// Liaison d'un résultat (docs/06 § 2)
{attribute 'pack_mode' := '1'}
TYPE ST_Bind :
STRUCT
    eTarget : E_BindTarget;
    nIndex : INT;
END_STRUCT
END_TYPE

(* stored: Version 1.1.0.1, ProductVersion 3.1.4024.12
   DUT ST_Bind: Id {044e01d3-6eb0-51b4-8a2a-b1068d56eaac} *)
